VAR_GLOBAL
    LinkData : ST_VC_LinkData;   // one per VisionCore connection, ~80 KB
END_VAR

(* stored: Version 1.1.0.1, ProductVersion 3.1.4024.12
   GVL GVL_VC: Id {116fb519-5010-436a-8702-082f9d29e6eb} *)
